Staubli VAL3: setIOvisible.pgx

public program setIOvisible(num x_nType)
  local string l_sbtn
  local num l_i
  local string l_slabel
  local num l_nSize
  local string l_slbl
  local string l_slbl1
  local string l_slbl2
  local num l_nSize1
begin
  call getSize(l_nSize,l_nSize1)
  switch x_nType
    case 0,1
      for l_i = 0 to 15
        l_slbl="lbl"+toString("",40+l_i)
        userPageSet("IO",l_slbl,"style.visibility","hidden")
      endFor
      for l_i = 0 to l_nSize-1
        l_slbl="lbl"+toString("",l_i)
        l_slbl1="lbl"+toString("",20+l_i)
        l_slbl2="btn"+toString("",60+l_i)
        userPageSet("IO",l_slbl,"style.visibility","visible")
        userPageSet("IO",l_slbl1,"style.visibility","visible")
        userPageSet("IO",l_slbl2,"style.visibility","visible")
      endFor
      if l_nSize<16
        for l_i = l_nSize to 15
          l_slbl="lbl"+toString("",l_i)
          l_slbl1="lbl"+toString("",20+l_i)
          l_slbl2="btn"+toString("",60+l_i)
          userPageSet("IO",l_slbl,"style.visibility","hidden")
          userPageSet("IO",l_slbl1,"style.visibility","hidden")
          userPageSet("IO",l_slbl2,"style.visibility","hidden")
        endFor
      endIf
    break
    case 2,3
      for l_i = 0 to 15
        l_slbl="btn"+toString("",60+l_i)
        userPageSet("IO",l_slbl,"style.visibility","hidden")
      endFor
      for l_i = 0 to l_nSize1-1
        l_slbl="lbl"+toString("",l_i)
        l_slbl1="lbl"+toString("",20+l_i)
        l_slbl2="lbl"+toString("",40+l_i)
        userPageSet("IO",l_slbl,"style.visibility","visible")
        userPageSet("IO",l_slbl1,"style.visibility","visible")
        userPageSet("IO",l_slbl2,"style.visibility","visible")
      endFor
      if l_nSize1<16
        for l_i = l_nSize1 to 15
          l_slbl="lbl"+toString("",l_i)
          l_slbl1="lbl"+toString("",20+l_i)
          l_slbl2="lbl"+toString("",40+l_i)
          userPageSet("IO",l_slbl,"style.visibility","hidden")
          userPageSet("IO",l_slbl1,"style.visibility","hidden")
          userPageSet("IO",l_slbl2,"style.visibility","hidden")
        endFor
      endIf
    break
  endSwitch
end
